(* IEC 61131-3 sources: sis-interlock-demo/tests/POUs/Suites/FB_SisUnit_Test, 7 files *)

(* ---- DisabledCauseVotingNotCalled.method.decl.st ---- *)
// Выключенная причина: группа голосования не вызывается (состояние по умолчанию, событий группы
// нет), требования нет, следствие 2 под напряжением
METHOD PRIVATE DisabledCauseVotingNotCalled
VAR
    fbRig : FB_UnitRig;   // стенд
END_VAR

(* ---- EventsVotingBeforeCem.method.decl.st ---- *)
// В одном вызове события групп голосования идут раньше событий матрицы: ChannelInvalid группы 1,
// затем CauseDemand причины 1 (недостоверный канал 1oo2 VoteTrip даёт требование)
METHOD PRIVATE EventsVotingBeforeCem
VAR
    fbRig : FB_UnitRig;     // стенд
    stEv  : ST_SisEvent;    // событие
END_VAR

(* ---- ExternalCauseUsesExtDemand.method.decl.st ---- *)
// Причина с источником External берёт требование из xExtDemand без голосования: фиксация, следствие 2
// обесточено, состояние группы — значения по умолчанию
METHOD PRIVATE ExternalCauseUsesExtDemand
VAR
    fbRig : FB_UnitRig;   // стенд
END_VAR

(* ---- Setup.method.decl.st ---- *)
// Стенд узла: 3 причины, 2 следствия, без срабатывания при старте.
//   1 — голосование DI 1oo2 (VoteTrip, байпас до 10 с), задержка 2 с;
//   2 — внешняя (xExtDemand), без задержки;
//   3 — выключена (группа DI 1oo1 задана).
//   Следствие 1 — причина 1 (16#0001); 2 — причины 2, 3 (16#0006). Каналы групп 1 и 3 — в норме.
METHOD Setup
VAR_IN_OUT
    fbRig : FB_UnitRig;    // стенд
END_VAR
VAR
    stCem  : ST_CemCfg;    // матрица
    stVote : ST_VotingCfg; // группа голосования
    uiK    : UINT;         // номер канала
END_VAR

(* ---- Setup.method.impl.st ---- *)
stCem.uiCauseCount := 3;
stCem.uiEffectCount := 2;
stCem.xStartTripped := FALSE;
stCem.astCause[1].xEnable := TRUE;
stCem.astCause[1].eSource := E_CauseSource.Voting;
stCem.astCause[1].tDelay := T#2S;
stCem.astCause[2].xEnable := TRUE;
stCem.astCause[2].eSource := E_CauseSource.External;
stCem.astCause[3].xEnable := FALSE;
stCem.astCause[3].eSource := E_CauseSource.Voting;
stCem.astEffect[1].eSafeState := E_SafeState.Closed;
stCem.astEffect[1].wCauseMask := 16#0001;
stCem.astEffect[2].eSafeState := E_SafeState.Stopped;
stCem.astEffect[2].wCauseMask := 16#0006;
stCem.wMatrixCrc := F_CemCrc(stCfg := stCem);
fbRig.stCemCfg := stCem;

stVote.eArch := E_VoteArch.Vote1oo2;
stVote.ePolicy := E_DegradePolicy.VoteTrip;
stVote.eInput := E_SisInputKind.Discrete;
stVote.xDiHealthy := TRUE;
stVote.tBypassMax := T#10S;
stVote.uiMaxBypass := 1;
fbRig.astVoteCfg[1] := stVote;
stVote.eArch := E_VoteArch.Vote1oo1;
stVote.uiMaxBypass := 0;
fbRig.astVoteCfg[3] := stVote;

FOR uiK := 1 TO GVL_Const.SIS_VOTE_CH_MAX DO
    fbRig.astIn[1].axDi[uiK] := TRUE;
    fbRig.astIn[1].axDiValid[uiK] := TRUE;
    fbRig.astIn[3].axDi[uiK] := TRUE;
    fbRig.astIn[3].axDiValid[uiK] := TRUE;
END_FOR

(* ---- TimeSourcePassedToChildren.method.decl.st ---- *)
// Источник времени узла передаётся группам и матрице: байпас группы 1 истекает ровно через 10 с
// подменного времени, задержка причины — ровно через 2 с
METHOD PRIVATE TimeSourcePassedToChildren
VAR
    fbRig : FB_UnitRig;   // стенд
END_VAR

(* ---- VotingCfgErrorTripsOnlyThatCause.method.decl.st ---- *)
// Ошибка конфигурации группы 1 — требование только причины 1: она срабатывает через обычную задержку
// 2 с, следствие 2 и причина 2 работают как обычно
METHOD PRIVATE VotingCfgErrorTripsOnlyThatCause
VAR
    fbRig : FB_UnitRig;     // стенд
    stDef : ST_VotingCfg;   // конфигурация по умолчанию (ошибка)
END_VAR
